TYPE E_NC_State :
(
	E_NC_State_INIT := 0,
	E_NC_State_IDLE := 1,
	E_NC_State_RUN := 7,
	E_NC_State_ABORT := 8,
	E_NC_State_ERROR := 9
);
END_TYPE

(* stored: Version 1.1.0.1, ProductVersion 3.1.4024.9
   DUT E_NC_State: Id {3a7dfb51-5f9b-40d0-b4df-f2633044854d} *)
